{attribute 'qualified_only'}
{attribute 'strict'}
TYPE E_CtlMd : 
(
	e_1 := 1, (*local*)
	e_2 := 2, (*remote*)
	e_3 := 3, (*auto*)
	e_4 := 4 (*test*)
) SINT;
END_TYPE

(* stored: Version 1.1.0.1
   DUT E_CtlMd: Id {3b27b253-7721-44f7-a2ed-bee8e6aa99b7} *)
